(* IEC 61131-3 sources: Test-Git_ESME26/TestProgettoESME_26.fbsproj/PacDriveLib Migration/Motion/Homing/PDL_FB_HomeIn.fb.st^, 4 files *)

(* ---- InitInterfaces.meth.st ---- *)
METHOD PRIVATE InitInterfaces : BOOL
VAR_INPUT
END_VAR

VAR
	ifGetParentDevice      : DTSI.IF_GetParentDevice;
	ifDeviceAccess         : DTSI.IF_DeviceAccess;
END_VAR

InitInterfaces := FALSE;
IF i_ifDrive = 0 THEN
	SetDiagOutput(	i_etDiag	:= GD.ET_Diag.InputParameterInvalid,
					i_etDiagExt := PDL_ET_DiagExt.DriveInvalid,
					i_sMsg		:= 'i_ifDrive - Invalid Interface');
	RETURN;
ELSE
	xSuccess := __QUERYINTERFACE(i_ifDrive, ifGetParentDevice);
	IF NOT xSuccess OR ifGetParentDevice = 0 THEN
		SetDiagOutput(	i_etDiag	:= GD.ET_Diag.InputParameterInvalid,
						i_etDiagExt := PDL_ET_DiagExt.DriveInvalid,
						i_sMsg		:= 'i_ifDrive - IF_GetParentDevice not implemented.');
		RETURN;
	END_IF
	ifDeviceAccess := ifGetParentDevice.GetParentDevice();

	xSuccess := __QUERYINTERFACE(ifDeviceAccess,ifDriveConfigAccess );
	IF (NOT xSuccess OR ifDriveConfigAccess = 0) THEN
		SetDiagOutput(	i_etDiag	:= GD.ET_Diag.InputParameterInvalid,
						i_etDiagExt := PDL_ET_DiagExt.DriveInvalid,
						i_sMsg		:= 'i_ifDrive - IF_DriveConfig not implemented.');
		diState := 0;
		RETURN;
	END_IF
	ifDriveConfig := ifDriveConfigAccess.DriveConfig;

	xSuccess := __QUERYINTERFACE(ifDeviceAccess, ifDeviceTreeObjectAccess);
	IF xSuccess THEN
		sDriveName := ifDeviceTreeObjectAccess.DeviceTreeObject.Name;
	ELSE
		sDriveName := 'Axis';
	END_IF

	THIS^.fbHalt.Axis         := i_ifDrive;
	THIS^.fbStop.Axis         := i_ifDrive;
	THIS^.fbSetPos.Axis       := i_ifDrive;
	THIS^.fbMoveRelative.Axis := i_ifDrive;
END_IF

InitInterfaces := TRUE;

(* ---- InputParameterCheck.meth.st ---- *)
METHOD PRIVATE InputParameterCheck : BOOL
VAR_INPUT
END_VAR
VAR
	lrMaxAcc	: LREAL := 0;
	lrMaxVel	: LREAL := 0;
END_VAR

InputParameterCheck := FALSE;

lrMaxAcc := ifDriveConfig.MaxAcc;
lrMaxVel := ifDriveConfig.MaxVel;

IF (i_lrMaxTravel <= 0.0) THEN
	SetDiagOutput(i_etDiag := GD.ET_Diag.InputParameterInvalid, i_etDiagExt := PDL_ET_DiagExt.MaxTravelRange, i_sMsg := '0.0 < i_lrMaxTravel');
	RETURN;

ELSIF i_lrVel <= 0.0 OR (i_lrVel > lrMaxVel AND lrMaxVel <> 0) THEN
	SetDiagOutput(
		i_etDiag    := GD.ET_Diag.InputParameterInvalid,
		i_etDiagExt := PDL_ET_DiagExt.VelRange,
		i_sMsg      := STANDARD.CONCAT('0.0 < i_lrVel <= ', TO_STRING(lrMaxVel))
	);
	RETURN;

ELSIF (i_lrAcc <= 0.0 OR i_lrAcc > lrMaxAcc AND lrMaxAcc <> 0) THEN
	SetDiagOutput(
		i_etDiag    := GD.ET_Diag.InputParameterInvalid,
		i_etDiagExt := PDL_ET_DiagExt.AccRange,
		i_sMsg      := STANDARD.CONCAT('0.0 < i_lrAcc <= ', TO_STRING(lrMaxAcc))
	);
	RETURN;

ELSIF (i_lrDec <= 0.0 OR i_lrDec > lrMaxAcc AND lrMaxAcc <> 0) THEN
	SetDiagOutput(
		i_etDiag    := GD.ET_Diag.InputParameterInvalid,
		i_etDiagExt := PDL_ET_DiagExt.DecRange,
		i_sMsg      := STANDARD.CONCAT('0.0 < i_lrDec <= ', TO_STRING(lrMaxAcc))
	);
	RETURN;

ELSIF i_lrJerk <= 0.0 THEN
	SetDiagOutput(i_etDiag := GD.ET_Diag.InputParameterInvalid, i_etDiagExt := PDL_ET_DiagExt.JerkRange, i_sMsg := '0.0 < i_lrJerk');
	RETURN;
END_IF

THIS^.fbMoveRelative.Velocity     := i_lrVel;
THIS^.fbMoveRelative.Acceleration := i_lrAcc;
THIS^.fbMoveRelative.Deceleration := i_lrDec;
THIS^.fbMoveRelative.Jerk         := i_lrJerk;
THIS^.fbMoveRelative.BufferMode   := PLCO.MC_Buffer_Mode.Aborting;

THIS^.fbHalt.Jerk         := i_lrJerk;
THIS^.fbHalt.Deceleration := i_lrDec;
THIS^.fbHalt.BufferMode   := PLCO.MC_Buffer_Mode.Aborting;

THIS^.fbStop.Jerk         := i_lrJerk;
THIS^.fbStop.Deceleration := i_lrDec;

InputParameterCheck := TRUE;

(* ---- RegisterLoggerPoint.meth.st ---- *)
METHOD PUBLIC RegisterLoggerPoint
VAR_INPUT
	i_ifParent		: APL.IF_LoggerPoint;
	i_sName			: STRING[80];
END_VAR
VAR_OUTPUT
	q_etDiag		: GD.ET_Diag := GD.ET_Diag.Ok;
	q_etDiagExt		: PDL_ET_DiagExt := PDL_ET_DiagExt.Ok;
END_VAR
VAR
	etDiagBuffer		: GD.ET_Diag;
	etDiagExtBufferAPL	: APL.ET_DiagExt;
END_VAR

THIS^.fbLoggerPoint.RegisterLoggerPoint(	i_ifParent		:= i_ifParent,
											i_sName			:= i_sName,
											i_sType			:= 'FB_HomeIn',
											i_sSource		:= 'PDL',
											q_etDiag		=> etDiagBuffer,
											q_etDiagExt		=> etDiagExtBufferAPL);
IF (etDiagBuffer <> GD.ET_Diag.Ok) THEN
	CASE etDiagExtBufferAPL OF
		APL.ET_DiagExt.ParentInvalid:
			q_etDiag := GD.ET_Diag.InputParameterInvalid;
			q_etDiagExt := PDL_ET_DiagExt.ParentInvalid;

		APL.ET_DiagExt.ParentNotRegistered:
			q_etDiag := GD.ET_Diag.InputParameterInvalid;
			q_etDiagExt := PDL_ET_DiagExt.ParentNotRegistered;

		APL.ET_DiagExt.MaxNumberOfLoggerPointsExeeded:
			q_etDiag := GD.ET_Diag.InputParameterInvalid;
			q_etDiagExt := PDL_ET_DiagExt.MaxNumberOfLoggerPointsExeeded;

	ELSE
		q_etDiag := GD.ET_Diag.UnexpectedProgramBehavior;
		q_etdiagExt := PDL_ET_DiagExt.UnexpectedDiagExt;
	END_CASE
END_IF

(* ---- SetDiagOutput.meth.st ---- *)
METHOD PRIVATE SetDiagOutput : BOOL
VAR_INPUT
	i_etDiag	: GD.ET_Diag;
	i_etDiagExt	: PDL_ET_DiagExt;
	i_sMsg		: STRING[80];
END_VAR

IF i_etDiag <> GD.ET_Diag.Ok THEN
	q_xReady := FALSE;
END_IF
IF q_etDiag = GD.ET_Diag.OK OR i_etDiagExt = PDL_ET_DiagExt.Disabled THEN
	q_etDiag := i_etDiag;
	q_etDiagExt := i_etDiagExt;
	q_sMsg := i_sMsg;

	IF(i_etDiag = GD.ET_Diag.Ok) AND (THIS^.fbLoggerPoint.etLogLevel >= APL.ET_LogLevel.StatusMessage) THEN
		THIS^.fbLoggerPoint.AddLogEntry(	i_etLogLevel	:= APL.ET_LogLevel.StatusMessage,
											i_etDiag		:= q_etDiag,
											i_udiDiagExt	:= q_etDiagExt,
											i_sMessage		:= SE_CTBX.FC_MultiConcat(	i_sString1	:= Standard.CONCAT('ET_Diag: ', GD.FC_EtDiagToString(q_etDiag)),
																				i_sString2	:= Standard.CONCAT(' PDL_ET_DiagExt: ', PDL_FC_EtDiagExtToString(q_etDiagExt)),
																				i_sString3	:= Standard.CONCAT(' sMsg: ', q_sMsg),
																				i_sString4	:= ''),
											q_etDiag		:= ,	// ignore result
											q_etDiagExt		:= );	// ignore result
	ELSIF(i_etDiag = GD.ET_Diag.UnexpectedProgramBehavior) AND (THIS^.fbLoggerPoint.etLogLevel >= APL.ET_LogLevel.CriticalException) THEN
		THIS^.fbLoggerPoint.AddLogEntry(	i_etLogLevel	:= APL.ET_LogLevel.CriticalException,
											i_etDiag		:= q_etDiag,
											i_udiDiagExt	:= q_etDiagExt,
											i_sMessage		:= SE_CTBX.FC_MultiConcat(	i_sString1	:= Standard.CONCAT('ET_Diag: ', GD.FC_EtDiagToString(q_etDiag)),
																				i_sString2	:= Standard.CONCAT(' PDL_ET_DiagExt: ', PDL_FC_EtDiagExtToString(q_etDiagExt)),
																				i_sString3	:= Standard.CONCAT(' sMsg: ', q_sMsg),
																				i_sString4	:= ''),
											q_etDiag		:= ,	// ignore result
											q_etDiagExt		:= );	// ignore result
	ELSIF(i_etDiag <> GD.ET_Diag.Ok) AND (THIS^.fbLoggerPoint.etLogLevel >= APL.ET_LogLevel.Exception) THEN
		THIS^.fbLoggerPoint.AddLogEntry(	i_etLogLevel	:= APL.ET_LogLevel.Exception,
											i_etDiag		:= q_etDiag,
											i_udiDiagExt	:= q_etDiagExt,
											i_sMessage		:= SE_CTBX.FC_MultiConcat(	i_sString1	:= Standard.CONCAT('ET_Diag: ', GD.FC_EtDiagToString(q_etDiag)),
																				i_sString2	:= Standard.CONCAT(' PDL_ET_DiagExt: ', PDL_FC_EtDiagExtToString(q_etDiagExt)),
																				i_sString3	:= Standard.CONCAT(' sMsg: ', q_sMsg),
																				i_sString4	:= ''),
											q_etDiag		:= ,	// ignore result
											q_etDiagExt		:= );	// ignore result
	END_IF
END_IF
